Fanuc KAREL source: kt00300.KL

-- PROVISIONAL review KL for V1013-1; original PC SHA256 54b6031b8ad978631b652bc563ec19507b5484cce66896dc9fbb5042189d2e3c
-- Incomplete behavior may be omitted. Consult companion uncertainty JSON. Do not deploy.
PROGRAM KT00300
%NOLOCKGROUP
VAR
  R1 : REAL
  OUT : BOOLEAN
-- UNRESOLVED_DECL H2 type=002017
BEGIN
  -- UNRESOLVED_PC offsets 5-16; opcodes 2E,23
  -- UNRESOLVED_PC offsets 21-35; opcodes 2E,22,9D,33,B4
  -- UNRESOLVED_PC offsets 40-63; opcodes 21,22,9D,33,B3,64,6E,23
  -- UNRESOLVED_PC offsets 68-72; opcodes 7F
END KT00300
